ABB RAPID module: ManyMoves.mod

MODULE MainModule
GLOBAL VAR robtarget robpoint0= p:{{-640.584, 506.980, 371.534},{0.374108, 0.285846, 0.853660, -0.222712}}{cfg 0,0,0,0}{EJ 0.000000000,0.000000000,0.000000000,0.000000000,0.000000000,0.000000000}
GLOBAL VAR robtarget robpoint1= p:{{-638.084, 504.480, 372.034},{0.374108, 0.285846, 0.853660, -0.222712}}{cfg 0,0,0,0}{EJ 0.000000000,0.000000000,0.000000000,0.000000000,0.000000000,0.000000000}
GLOBAL VAR robtarget robpoint2= p:{{-630.584, 496.980, 373.534},{0.374108, 0.285846, 0.853660, -0.222712}}{cfg 0,0,0,0}{EJ 0.000000000,0.000000000,0.000000000,0.000000000,0.000000000,0.000000000}
GLOBAL VAR robtarget robpoint3= p:{{-628.084, 494.480, 374.034},{0.374108, 0.285846, 0.853660, -0.222712}}{cfg 0,0,0,0}{EJ 0.000000000,0.000000000,0.000000000,0.000000000,0.000000000,0.000000000}
GLOBAL VAR robtarget robpoint4= p:{{-620.584, 486.980, 375.534},{0.374108, 0.285846, 0.853660, -0.222712}}{cfg 0,0,0,0}{EJ 0.000000000,0.000000000,0.000000000,0.000000000,0.000000000,0.000000000}
GLOBAL VAR robtarget robpoint5= p:{{-618.084, 484.480, 376.034},{0.374108, 0.285846, 0.853660, -0.222712}}{cfg 0,0,0,0}{EJ 0.000000000,0.000000000,0.000000000,0.000000000,0.000000000,0.000000000}
GLOBAL VAR robtarget robpoint6= p:{{-610.584, 476.980, 377.534},{0.374108, 0.285846, 0.853660, -0.222712}}{cfg 0,0,0,0}{EJ 0.000000000,0.000000000,0.000000000,0.000000000,0.000000000,0.000000000}
GLOBAL VAR robtarget robpoint7= p:{{-608.084, 474.480, 378.034},{0.374108, 0.285846, 0.853660, -0.222712}}{cfg 0,0,0,0}{EJ 0.000000000,0.000000000,0.000000000,0.000000000,0.000000000,0.000000000}
GLOBAL VAR robtarget robpoint8= p:{{-600.584, 466.980, 379.534},{0.374108, 0.285846, 0.853660, -0.222712}}{cfg 0,0,0,0}{EJ 0.000000000,0.000000000,0.000000000,0.000000000,0.000000000,0.000000000}
GLOBAL VAR robtarget robpoint9= p:{{-598.084, 464.480, 380.034},{0.374108, 0.285846, 0.853660, -0.222712}}{cfg 0,0,0,0}{EJ 0.000000000,0.000000000,0.000000000,0.000000000,0.000000000,0.000000000}
GLOBAL VAR robtarget robpoint10= p:{{-590.584, 456.980, 381.534},{0.374108, 0.285846, 0.853660, -0.222712}}{cfg 0,0,0,0}{EJ 0.000000000,0.000000000,0.000000000,0.000000000,0.000000000,0.000000000}
GLOBAL VAR robtarget robpoint11= p:{{-588.084, 454.480, 382.034},{0.374108, 0.285846, 0.853660, -0.222712}}{cfg 0,0,0,0}{EJ 0.000000000,0.000000000,0.000000000,0.000000000,0.000000000,0.000000000}
GLOBAL VAR robtarget robpoint12= p:{{-580.584, 446.980, 383.534},{0.374108, 0.285846, 0.853660, -0.222712}}{cfg 0,0,0,0}{EJ 0.000000000,0.000000000,0.000000000,0.000000000,0.000000000,0.000000000}
GLOBAL VAR robtarget robpoint13= p:{{-578.084, 444.480, 384.034},{0.374108, 0.285846, 0.853660, -0.222712}}{cfg 0,0,0,0}{EJ 0.000000000,0.000000000,0.000000000,0.000000000,0.000000000,0.000000000}
GLOBAL VAR robtarget robpoint14= p:{{-570.584, 436.980, 385.534},{0.374108, 0.285846, 0.853660, -0.222712}}{cfg 0,0,0,0}{EJ 0.000000000,0.000000000,0.000000000,0.000000000,0.000000000,0.000000000}
GLOBAL VAR robtarget robpoint15= p:{{-568.084, 434.480, 386.034},{0.374108, 0.285846, 0.853660, -0.222712}}{cfg 0,0,0,0}{EJ 0.000000000,0.000000000,0.000000000,0.000000000,0.000000000,0.000000000}
GLOBAL VAR robtarget robpoint16= p:{{-560.584, 426.980, 387.534},{0.374108, 0.285846, 0.853660, -0.222712}}{cfg 0,0,0,0}{EJ 0.000000000,0.000000000,0.000000000,0.000000000,0.000000000,0.000000000}
GLOBAL VAR robtarget robpoint17= p:{{-558.084, 424.480, 388.034},{0.374108, 0.285846, 0.853660, -0.222712}}{cfg 0,0,0,0}{EJ 0.000000000,0.000000000,0.000000000,0.000000000,0.000000000,0.000000000}
GLOBAL VAR robtarget robpoint18= p:{{-550.584, 416.980, 389.534},{0.374108, 0.285846, 0.853660, -0.222712}}{cfg 0,0,0,0}{EJ 0.000000000,0.000000000,0.000000000,0.000000000,0.000000000,0.000000000}
GLOBAL VAR robtarget robpoint19= p:{{-548.084, 414.480, 390.034},{0.374108, 0.285846, 0.853660, -0.222712}}{cfg 0,0,0,0}{EJ 0.000000000,0.000000000,0.000000000,0.000000000,0.000000000,0.000000000}

GLOBAL Proc main()
    wobj16.x = 1234.57
    wobj16.y = -98.765
    wobj16.z = 50.500
    wobj16.q1 = 0.965926
    wobj16.q2 = 0.000000
    wobj16.q3 = 0.000000
    wobj16.q4 = 0.258819
    tool03.x = 10.000
    tool03.y = 20.000
    tool03.z = 150.000
    tool03.q1 = 1.000000
    tool03.q2 = 0.000000
    tool03.q3 = 0.000000
    tool03.q4 = 0.000000
    MoveJ robpoint0,v500,z50,tool03,wobj16
    MoveL robpoint1,v500,z50,tool03,wobj16
    MoveJ robpoint2,v500,z50,tool03,wobj16
    MoveL robpoint3,v500,z50,tool03,wobj16
    MoveJ robpoint4,v500,z50,tool03,wobj16
    MoveL robpoint5,v500,z50,tool03,wobj16
    MoveJ robpoint6,v500,z50,tool03,wobj16
    MoveL robpoint7,v500,z50,tool03,wobj16
    MoveJ robpoint8,v500,z50,tool03,wobj16
    MoveL robpoint9,v500,z50,tool03,wobj16
    MoveJ robpoint10,v500,z50,tool03,wobj16
    MoveL robpoint11,v500,z50,tool03,wobj16
    MoveJ robpoint12,v500,z50,tool03,wobj16
    MoveL robpoint13,v500,z50,tool03,wobj16
    MoveJ robpoint14,v500,z50,tool03,wobj16
    MoveL robpoint15,v500,z50,tool03,wobj16
    MoveJ robpoint16,v500,z50,tool03,wobj16
    MoveL robpoint17,v500,z50,tool03,wobj16
    MoveJ robpoint18,v500,z50,tool03,wobj16
    MoveL robpoint19,v500,z50,tool03,wobj16
EndProc
EndModule
